Fanuc KAREL source: kd00023.KL

-- PROVISIONAL review KL for V940-1; original PC SHA256 d0ad9514288a18bdf430dca59206007df7a418aeeddadbc7b20c7d077d13af26
-- Incomplete behavior may be omitted. Consult companion uncertainty JSON. Do not deploy.
PROGRAM KD00023
%NOLOCKGROUP
VAR
  I : INTEGER
  J : INTEGER
  B : BOOLEAN
  R : REAL
  S : STRING[80]
  SAVED : INTEGER
BEGIN
  -- V9_ZERO_TABLE_METADATA_HINT layout=0001; no indexed target words; source/name/runtime held
  -- UNRESOLVED_PC offsets 5-17; opcodes 21,23
  -- UNRESOLVED_PC offsets 22-26; opcodes 7F
END KD00023
